Staubli VAL3: start.pgx

public program start()
begin
  // Program MAIN_1 start
  // Program generated by RoboDK v5.6.9 for RoboDK Industrial on 26/02/2024 09:58:20
  // Using nominal kinematics.
  nTraj=movej(jJoint[0],flange[0],mNomSpeed)
  nTraj=movej(jJoint[1],flange[0],mNomSpeed)
  nTraj=movel(pPoint[0],flange[0],mNomSpeed)
  do5=true
  do5=true
  do5=0.5
  do5=true
  do5=true
  do5=true
  do5=0.5
  do5=true
  var=val
  var=val
  WAIT FOR di5==true
  WAIT FOR di5==true
  WAIT FOR di5==0.5
  WAIT FOR di5==true
  WAIT FOR di5==true TIMEOUT=100.0
  WAIT FOR var==val
  WAIT FOR var==val TIMEOUT=100.0
  popUpMsg("Message")
  //call prog:REMOTE_PROG_CALL_171()
  CODE_INSERT_172
  // Insert Comment
  nTraj=movej(jJoint[2],tCad[0],mNomSpeed)
  nTraj=movel(pPoint[1],tCad[0],mSpeed[0])
  do5=true
  //call prog:PICK_PART_111()
  // Linear movement using joint targets is not supported. Change the target type to cartesian or use a joint movement.
  nTraj=movel(pPoint[2],tCad[0],mSpeed[1])
  // MoveSearch command not implemented
  nTraj=movel(pPoint[3],tCad[0],mSpeed[2])
  do5=false
  //call prog:PLACE_PART_112()
  nTraj=movel(pPoint[4],tCad[0],mSpeed[2])
  nTraj=movej(jJoint[3],tCad[0],mSpeed[3])
  nTraj=movec(pPoint[5],pPoint[6],tCad[0],mSpeed[3])
  // Circular movement using joint targets is not supported. Change the target type to cartesian or use a joint movement.
  nTraj=movel(pPoint[7],tCad[0],mSpeed[4])
  nTraj=movej(jJoint[4],tCad[0],mSpeed[4])
  // Warning: This post processor supports one reference frame only. Please use the Staubli VAL3 simplified post processor instead. Errors might follow.
  nTraj=movej(jJoint[5],tCad[0],mSpeed[4])
  nTraj=movel(pPoint[8],tCad[0],mSpeed[4])
  nTraj=movel(pPoint[9],tCad[0],mSpeed[4])
  nTraj=movel(pPoint[10],tCad[0],mSpeed[4])
  nTraj=movel(pPoint[11],tCad[0],mSpeed[4])
  nTraj=movel(pPoint[12],tCad[0],mSpeed[4])
  nTraj=movel(pPoint[13],tCad[0],mSpeed[4])
  nTraj=movel(pPoint[14],tCad[0],mSpeed[4])
  nTraj=movej(jJoint[6],tCad[0],mSpeed[4])
  //call prog:EVENT_PROG_START_101()
  // Warning: This post processor supports one reference frame only. Please use the Staubli VAL3 simplified post processor instead. Errors might follow.
  // Show Tool 1
  nTraj=movej(jJoint[7],tCad[0],mSpeed[5])
  //call prog:EVENT_PATH_APPROACH_102()
  nTraj=movel(pPoint[15],tCad[0],mSpeed[5])
  nTraj=movel(pPoint[16],tCad[0],mSpeed[5])
  //call prog:EVENT_PATH_START_103()
  nTraj=movel(pPoint[17],tCad[0],mSpeed[6])
  nTraj=movel(pPoint[18],tCad[0],mSpeed[6])
  nTraj=movel(pPoint[19],tCad[0],mSpeed[6])
  nTraj=movel(pPoint[20],tCad[0],mSpeed[6])
  nTraj=movel(pPoint[21],tCad[0],mSpeed[6])
  nTraj=movel(pPoint[22],tCad[0],mSpeed[6])
  nTraj=movel(pPoint[23],tCad[0],mSpeed[6])
  nTraj=movel(pPoint[24],tCad[0],mSpeed[6])
  nTraj=movel(pPoint[25],tCad[0],mSpeed[6])
  nTraj=movel(pPoint[26],tCad[0],mSpeed[6])
  nTraj=movel(pPoint[27],tCad[0],mSpeed[6])
  nTraj=movel(pPoint[28],tCad[0],mSpeed[6])
  nTraj=movel(pPoint[29],tCad[0],mSpeed[6])
  nTraj=movel(pPoint[30],tCad[0],mSpeed[6])
  nTraj=movel(pPoint[31],tCad[0],mSpeed[6])
  nTraj=movel(pPoint[32],tCad[0],mSpeed[6])
  nTraj=movel(pPoint[33],tCad[0],mSpeed[6])
  nTraj=movel(pPoint[34],tCad[0],mSpeed[6])
  nTraj=movel(pPoint[35],tCad[0],mSpeed[6])
  nTraj=movel(pPoint[36],tCad[0],mSpeed[6])
  nTraj=movel(pPoint[37],tCad[0],mSpeed[6])
  nTraj=movel(pPoint[38],tCad[0],mSpeed[6])
  nTraj=movel(pPoint[39],tCad[0],mSpeed[6])
  nTraj=movel(pPoint[40],tCad[0],mSpeed[6])
  nTraj=movel(pPoint[41],tCad[0],mSpeed[6])
  nTraj=movel(pPoint[42],tCad[0],mSpeed[6])
  nTraj=movel(pPoint[43],tCad[0],mSpeed[6])
  nTraj=movel(pPoint[44],tCad[0],mSpeed[6])
  nTraj=movel(pPoint[45],tCad[0],mSpeed[6])
  nTraj=movel(pPoint[46],tCad[0],mSpeed[6])
  nTraj=movel(pPoint[47],tCad[0],mSpeed[6])
  nTraj=movel(pPoint[48],tCad[0],mSpeed[6])
  nTraj=movel(pPoint[49],tCad[0],mSpeed[6])
  nTraj=movel(pPoint[50],tCad[0],mSpeed[6])
  nTraj=movel(pPoint[51],tCad[0],mSpeed[6])
  nTraj=movel(pPoint[52],tCad[0],mSpeed[6])
  nTraj=movel(pPoint[53],tCad[0],mSpeed[6])
  nTraj=movel(pPoint[54],tCad[0],mSpeed[6])
  nTraj=movel(pPoint[55],tCad[0],mSpeed[6])
  nTraj=movel(pPoint[56],tCad[0],mSpeed[6])
  nTraj=movel(pPoint[57],tCad[0],mSpeed[6])
  nTraj=movel(pPoint[58],tCad[0],mSpeed[6])
  nTraj=movel(pPoint[59],tCad[0],mSpeed[6])
  nTraj=movel(pPoint[60],tCad[0],mSpeed[6])
  nTraj=movel(pPoint[61],tCad[0],mSpeed[6])
  //call prog:EVENT_PATH_FINISH_105()
  nTraj=movel(pPoint[62],tCad[0],mSpeed[7])
  nTraj=movel(pPoint[63],tCad[0],mSpeed[7])
  //call prog:EVENT_PATH_RETRACT_106()
  //call prog:EVENT_PROG_FINISH_107()
  // Warning: This post processor supports one reference frame only. Please use the Staubli VAL3 simplified post processor instead. Errors might follow.
  nTraj=movej(jJoint[8],tCad[0],mSpeed[7])
  delay(1.250)
  nTraj=movel(pPoint[64],tCad[0],mSpeed[7])
  WAIT FOR di1==true
  nTraj=movel(pPoint[65],tCad[0],mSpeed[7])
  //call prog:PROG 1 _.-[]/\;,><&*:%=+@!#^|?^ with a very long name and special characters()

  waitEndMove()
  // Program MAIN_1 end
  // Program PROG1_withaverylongnameandspecialcharacters start
  // This is a subprogram call to PROG_1
  // Warning: This post processor supports one reference frame only. Please use the Staubli VAL3 simplified post processor instead. Errors might follow.
  nTraj=movej(jJoint[9],tCad[1],mSpeed[7])

  waitEndMove()
  // Program PROG1_withaverylongnameandspecialcharacters end

end
